{attribute 'qualified_only'}
{attribute 'strict'}
{attribute 'to_string'}
TYPE E_ValueType :
(
	E_String := 0,
	E_TraceId,
	E_SpanId,
	E_AnyValue,
	E_KeyValue,
	E_Number
);
END_TYPE

(* stored: Version 1.1.0.1
   EnumerationTextList E_ValueType: Id {2fd589b6-3af6-4d4c-9efd-75488ffbdda6} *)
